(* IEC 61131-3 sources: STAR-PLC-Agent/results/raw/codex_matrix_resume_20261114/codex_deepseek/SELF009/generation/compiler_records/compile_00, 1 file *)

(* ---- FB_Task.st ---- *)
FUNCTION_BLOCK FB_Task
VAR_INPUT
    PartPulse : BOOL;
    Reset : BOOL;
    Target : USINT;
END_VAR
VAR_OUTPUT
    Count : USINT := 0;
    Complete : BOOL := FALSE;
    Error : BOOL := FALSE;
END_VAR
VAR
    previous_pulse : BOOL := FALSE;
END_VAR

Error := (Target < 1) OR (Target > 20);

IF Error OR Reset THEN
    Count := 0;
    Complete := FALSE;
ELSE
    IF PartPulse AND NOT previous_pulse AND (Count < Target) THEN
        Count := Count + 1;
    ELSIF Count > Target THEN
        Count := Target;
    END_IF;
    Complete := (Count >= Target);
END_IF;

previous_pulse := PartPulse;
END_FUNCTION_BLOCK
